# B&R Automation Studio project AS_Project (part 2)

#### Convert.c - dbGetData data conversion
```c
/********************************************************************
 * Library: AltDB
 * File: Convert.c
 ********************************************************************
 * dbGetData data conversion (Section 11). Converts the raw column
 * value bytes stored by Token.c (gConn[slot].ColValue[columnIdx])
 * into one of the DB_SQL_* target layouts of Table 22.
 *
 * Scope: the full conversion matrix (Table 23) is implemented for
 * the practically important source/target combinations. Combinations
 * marked '-' in Table 23, and sources this library cannot decode at
 * all (SQL_VARIANT, XML, UDT), are rejected with dbERR_DATABASE /
 * SQLSTATE 07006, matching the "not allowed" semantics of the
 * specification. DATETIMEOFFSET is read as if it were DATETIME2 (the
 * trailing minute-offset field is ignored, i.e. treated as UTC/local
 * time) - a documented simplification, see Common.h.
 ********************************************************************/
#include <bur/plctypes.h>
#include <runtime.h>
#include <AsTCP.h>
#include <AltDB.h>
#include "Common.h"
#include <string.h>

enum {
	FAM_INT, FAM_FLOAT, FAM_DECIMAL, FAM_MONEY, FAM_CHAR, FAM_BINARY,
	FAM_DATE, FAM_TIME, FAM_DATETIME, FAM_DATETIME2, FAM_GUID, FAM_UNSUPPORTED
};

static int Family(unsigned char t)
{
	switch (t) {
	case 0x30: case 0x32: case 0x34: case 0x38: case 0x7F:
	case 0x26: case 0x68:
		return FAM_INT;
	case 0x3B: case 0x3E: case 0x6D:
		return FAM_FLOAT;
	case 0x6A: case 0x6C:
		return FAM_DECIMAL;
	case 0x3C: case 0x7A: case 0x6E:
		return FAM_MONEY;
	case 0xA7: case 0xAF: case 0xE7: case 0xEF:
	case 0x2F: case 0x27:
	case 0x23: case 0x63:
		return FAM_CHAR;
	case 0xA5: case 0xAD: case 0x2D: case 0x25: case 0x22:
		return FAM_BINARY;
	case 0x28:
		return FAM_DATE;
	case 0x29:
		return FAM_TIME;
	case 0x3A: case 0x3D: case 0x6F:
		return FAM_DATETIME;
	case 0x2A: case 0x2B:
		return FAM_DATETIME2;
	case 0x24:
		return FAM_GUID;
	default:
		return FAM_UNSUPPORTED;
	}
}

static long long ReadIntValue(const unsigned char *p, UDINT len)
{
	unsigned long long u = 0;
	UDINT i;
	for (i = 0; i < len && i < 8; i++) u |= ((unsigned long long)p[i]) << (8 * i);
	if (len == 1) return (long long)u;        /* tinyint/bit: unsigned */
	if (len == 2) return (long long)(short)(unsigned short)u;
	if (len == 4) return (long long)(DINT)(UDINT)u;
	return (long long)u;
}

static long long ReadMoneyValue(const unsigned char *p, UDINT len)
{
	if (len == 4) return (long long)(DINT)AltDB_ReadLE32(p);
	{
		DINT hi = (DINT)AltDB_ReadLE32(p);
		UDINT lo = AltDB_ReadLE32(p + 4);
		return ((long long)hi << 32) | (long long)lo;
	}
}

static double ReadFloatValue(const unsigned char *p, UDINT len)
{
	if (len == 4) {
		union { UDINT u; float f; } v;
		v.u = AltDB_ReadLE32(p);
		return (double)v.f;
	} else {
		union { unsigned long long u; double d; } v;
		v.u = AltDB_ReadLE64(p);
		return v.d;
	}
}

/* value = integer / 10^scale, formatted as a decimal string */
static UDINT FormatScaledI64(long long v, USINT scale, char *dst, UDINT dstCap)
{
	unsigned char mag[8];
	BOOL positive = (v >= 0);
	unsigned long long u = positive ? (unsigned long long)v : (unsigned long long)(-(v + 1)) + 1ULL;
	UDINT i;
	for (i = 0; i < 8; i++) { mag[i] = (unsigned char)(u & 0xFF); u >>= 8; }
	return AltDB_FormatDecimal(mag, 8, positive, scale, dst, dstCap);
}

/* Decodes a DECIMALN/NUMERICN value (1 sign byte + little-endian
 * magnitude) into a plain double; sufficient precision for REAL /
 * DOUBLE targets (exact string output uses AltDB_FormatDecimal
 * directly for the CHAR target). */
static double DecimalToDouble(const unsigned char *raw, UDINT len, USINT scale)
{
	double v = 0.0;
	UDINT magLen = (len > 0) ? len - 1 : 0;
	BOOL positive = (len > 0) ? (raw[0] != 0) : TRUE;
	double divisor = 1.0;
	UDINT i;

	for (i = magLen; i > 0; i--) {
		v = v * 256.0 + (double)raw[i];
	}
	if (!positive) v = -v;
	for (i = 0; i < scale; i++) divisor *= 10.0;
	return v / divisor;
}

static void WriteGuidString(const unsigned char *g, char *dst)
{
	static const char *hex = "0123456789ABCDEF";
	static const int order[16] = {3,2,1,0, 5,4, 7,6, 8,9, 10,11,12,13,14,15};
	int i, p = 0;
	for (i = 0; i < 16; i++) {
		unsigned char b = g[order[i]];
		dst[p++] = hex[(b >> 4) & 0xF];
		dst[p++] = hex[b & 0xF];
		if (i == 3 || i == 5 || i == 7 || i == 9) dst[p++] = '-';
	}
	dst[p] = 0;
}

/* ---------------- date / time decoding (Section 10.9) ---------------- */

/* Howard Hinnant's civil_from_days algorithm (public domain formula),
 * valid over the whole proleptic Gregorian calendar. z = days since
 * 1970-01-01. */
static void CivilFromDays(long long z, INT *y, UINT *m, UINT *d)
{
	long long era;
	unsigned doe, yoe, doy, mp;

	z += 719468;
	era = (z >= 0 ? z : z - 146096) / 146097;
	doe = (unsigned)(z - era * 146097);
	yoe = (doe - doe / 1460 + doe / 36524 - doe / 146096) / 365;
	doy = doe - (365 * yoe + yoe / 4 - yoe / 100);
	mp = (5 * doy + 2) / 153;
	*d = (UINT)(doy - (153 * mp + 2) / 5 + 1);
	*m = (UINT)(mp + (mp < 10 ? 3 : -9));
	*y = (INT)((long long)yoe + era * 400 + (*m <= 2 ? 1 : 0));
}

typedef struct { INT y; UINT mo; UINT d; UINT h; UINT mi; UINT s; UDINT frac; USINT fracDigits; } DecodedDT;

/* days-since-0001-01-01 -> civil date */
static void DateFromDbDays(UDINT dbDays, INT *y, UINT *m, UINT *d)
{
	/* days_from_civil(1,1,1) = -719162 (date 0001-01-01 relative to 1970-01-01) */
	CivilFromDays((long long)dbDays - 719162LL, y, m, d);
}

static BOOL DecodeDateTime(int fam, unsigned char dataType, const unsigned char *raw, UDINT rawLen, USINT scale, DecodedDT *out)
{
	memset(out, 0, sizeof(*out));

	if (fam == FAM_DATE) {
		UDINT days = raw[0] | ((UDINT)raw[1] << 8) | ((UDINT)raw[2] << 16);
		DateFromDbDays(days, &out->y, &out->mo, &out->d);
		return TRUE;
	}
	if (fam == FAM_TIME || fam == FAM_DATETIME2) {
		UDINT dateBytes = (fam == FAM_DATETIME2) ? 3 : 0;
		UDINT offsetBytes = (dataType == 0x2B) ? 2 : 0;
		UDINT timeLen = (rawLen > dateBytes + offsetBytes) ? rawLen - dateBytes - offsetBytes : rawLen;
		UDINT i;
		unsigned long long ticks = 0;
		unsigned long long divisor = 1;
		UDINT secTotal;

		for (i = 0; i < timeLen && i < 8; i++) ticks |= ((unsigned long long)raw[i]) << (8 * i);
		for (i = 0; i < scale; i++) divisor *= 10ULL;
		secTotal = (UDINT)(ticks / divisor);
		out->frac = (UDINT)(ticks % divisor);
		out->fracDigits = scale;
		out->h = secTotal / 3600; out->mi = (secTotal / 60) % 60; out->s = secTotal % 60;

		if (fam == FAM_DATETIME2) {
			UDINT days = raw[timeLen] | ((UDINT)raw[timeLen + 1] << 8) | ((UDINT)raw[timeLen + 2] << 16);
			DateFromDbDays(days, &out->y, &out->mo, &out->d);
		}
		return TRUE;
	}
	if (fam == FAM_DATETIME) {
		if (rawLen == 4) { /* SMALLDATETIME: days(2,u16) + minutes(2,u16) since 1900-01-01 */
			UINT days = (UINT)AltDB_ReadLE16(raw);
			UINT minutes = (UINT)AltDB_ReadLE16(&raw[2]);
			CivilFromDays((long long)days - 25567LL, &out->y, &out->mo, &out->d); /* 1900-01-01 vs 1970-01-01 */
			out->h = minutes / 60; out->mi = minutes % 60; out->s = 0;
		} else { /* DATETIME: days(4,signed) + ticks(4,u32) of 1/300s since midnight */
			DINT days = (DINT)AltDB_ReadLE32(raw);
			UDINT ticks = AltDB_ReadLE32(&raw[4]);
			UDINT secTotal = ticks / 300;
			CivilFromDays((long long)days - 25567LL, &out->y, &out->mo, &out->d);
			out->h = secTotal / 3600; out->mi = (secTotal / 60) % 60; out->s = secTotal % 60;
		}
		return TRUE;
	}
	return FALSE;
}

static UDINT FormatDateTimeChar(int fam, const DecodedDT *dt, char *dst, UDINT cap)
{
	UDINT n = 0;
	char tmp[16];
	UDINT tn;

#define APPEND_NUM(v, width) do { \
		UDINT k; tn = (UDINT)AltDB_FormatI64((v), tmp, sizeof(tmp)); \
		for (k = tn; k < (UDINT)(width); k++) { if (n < cap) dst[n++] = '0'; } \
		for (k = 0; k < tn; k++) { if (n < cap) dst[n++] = tmp[k]; } \
	} while (0)

	if (fam == FAM_DATE || fam == FAM_DATETIME || fam == FAM_DATETIME2) {
		APPEND_NUM(dt->y, 4);
		if (n < cap) dst[n++] = '-';
		APPEND_NUM((long long)dt->mo, 2);
		if (n < cap) dst[n++] = '-';
		APPEND_NUM((long long)dt->d, 2);
		if (fam == FAM_DATE) { if (n < cap) dst[n] = 0; return n; }
		if (n < cap) dst[n++] = ' ';
	}

	APPEND_NUM((long long)dt->h, 2);
	if (n < cap) dst[n++] = ':';
	APPEND_NUM((long long)dt->mi, 2);
	if (n < cap) dst[n++] = ':';
	APPEND_NUM((long long)dt->s, 2);
	if (dt->fracDigits > 0) {
		if (n < cap) dst[n++] = '.';
		APPEND_NUM((long long)dt->frac, dt->fracDigits);
	}
	if (n < cap) dst[n] = 0;
	return n;
#undef APPEND_NUM
}

static void PutCharResult(const char *text, UDINT textLen, UDINT pData, UDINT dataSize,
                           UINT *status, INT *dbError, UDINT *actDataSize)
{
	UDINT required = textLen + 1;
	if (dataSize < required) {
		*status = dbERR_BUFFER_SIZE; *dbError = DB_SQL_ERROR; *actDataSize = required;
		return;
	}
	memcpy((void *)pData, text, textLen);
	((char *)pData)[textLen] = 0;
	*status = ERR_OK; *dbError = 0; *actDataSize = required;
}

void AltDB_GetData(UDINT slot, UDINT columnIdx, INT dataType, UDINT pData, UDINT dataSize,
                      UINT *status, INT *dbError, UDINT *actDataSize)
{
	ConnSlot *c = &gConn[slot];
	UDINT idx;
	ColumnInfo *col;
	int fam;
	const unsigned char *raw;
	UDINT rawLen;

	*actDataSize = 0;

	if (!c->RowReady) { *status = dbERR_SQL_EXECUTE_REQUIRED; *dbError = DB_SQL_ERROR; return; }
	if (columnIdx == 0 || columnIdx > (UDINT)c->ColumnCount || columnIdx > ND_MAX_COLUMNS) {
		*status = dbERR_INVALID_COLUMN; *dbError = DB_SQL_ERROR; return;
	}
	if (pData == 0) { *status = dbERR_NULLPOINTER; *dbError = DB_SQL_ERROR; return; }

	idx = columnIdx - 1;
	if (c->ColAlreadyRead[idx]) { *status = dbERR_DATABASE; *dbError = DB_SQL_NO_DATA; return; }

	if (c->ColIsNull[idx]) {
		*status = ERR_OK; *dbError = 0; *actDataSize = 0xFFFFFFFFUL;
		c->ColAlreadyRead[idx] = TRUE;
		return;
	}

	col = &c->Columns[idx];
	raw = c->ColValue[idx];
	rawLen = c->ColValueLen[idx];
	if (rawLen > ND_MAX_COL_VALUE_LEN) rawLen = ND_MAX_COL_VALUE_LEN;

	if (!col->Supported) {
		AltDB_DiagPushClient(slot, "07006", "source column type is not convertible by this library");
		*status = dbERR_DATABASE; *dbError = DB_SQL_ERROR; return;
	}

	fam = Family(col->DataType);

	switch (dataType) {

	case 1: { /* DB_SQL_CHAR */
		char text[600];
		UDINT n = 0;

		switch (fam) {
		case FAM_CHAR:
			if (col->IsUnicode) n = AltDB_WireToConn(c->Encoding, raw, rawLen, (unsigned char *)text, sizeof(text) - 1);
			else { n = (rawLen < sizeof(text) - 1) ? rawLen : sizeof(text) - 1; memcpy(text, raw, n); }
			break;
		case FAM_BINARY: {
			static const char *hex = "0123456789ABCDEF";
			UDINT i;
			for (i = 0; i < rawLen && n + 2 < sizeof(text); i++) {
				text[n++] = hex[(raw[i] >> 4) & 0xF];
				text[n++] = hex[raw[i] & 0xF];
			}
			break;
		}
		case FAM_INT:
			n = (UDINT)AltDB_FormatI64(ReadIntValue(raw, rawLen), text, sizeof(text));
			break;
		case FAM_MONEY:
			n = FormatScaledI64(ReadMoneyValue(raw, rawLen), 4, text, sizeof(text));
			break;
		case FAM_DECIMAL:
			n = AltDB_FormatDecimal(&raw[1], (rawLen > 0) ? rawLen - 1 : 0, raw[0] != 0, col->Scale, text, sizeof(text));
			break;
		case FAM_FLOAT:
			n = AltDB_FormatDouble(ReadFloatValue(raw, rawLen), (rawLen == 4) ? 7 : 15, text, sizeof(text));
			break;
		case FAM_GUID:
			if (rawLen >= 16) { WriteGuidString(raw, text); n = (UDINT)strlen(text); }
			break;
		case FAM_DATE: case FAM_TIME: case FAM_DATETIME: case FAM_DATETIME2: {
			DecodedDT dt;
			if (DecodeDateTime(fam, col->DataType, raw, rawLen, col->Scale, &dt)) {
				n = FormatDateTimeChar(fam, &dt, text, sizeof(text));
			}
			break;
		}
		default:
			AltDB_DiagPushClient(slot, "07006", "source column type is not convertible to DB_SQL_CHAR");
			*status = dbERR_DATABASE; *dbError = DB_SQL_ERROR; return;
		}
		PutCharResult(text, n, pData, dataSize, status, dbError, actDataSize);
		if (*status == ERR_OK) c->ColAlreadyRead[idx] = TRUE;
		return;
	}

	case -6: case 5: case 4: case -25: { /* TINYINT / SMALLINT / INTEGER / BIGINT */
		long long v;
		UDINT needed = (dataType == -6) ? 1 : (dataType == 5) ? 2 : (dataType == 4) ? 4 : 8;

		if (fam == FAM_INT) v = ReadIntValue(raw, rawLen);
		else if (fam == FAM_MONEY) v = ReadMoneyValue(raw, rawLen) / 10000;
		else if (fam == FAM_DECIMAL) v = (long long)DecimalToDouble(raw, rawLen, col->Scale);
		else if (fam == FAM_FLOAT) v = (long long)ReadFloatValue(raw, rawLen);
		else {
			AltDB_DiagPushClient(slot, "07006", "source column type is not convertible to an integer type");
			*status = dbERR_DATABASE; *dbError = DB_SQL_ERROR; return;
		}
				/* AsDB compatibility: allow BIGINT -> UDINT */

		if (dataType == -25 && dataSize == 4)
		{
			UDINT tmp = (UDINT)v;
			memcpy((void *)pData, &tmp, 4);
			*status = ERR_OK;
			*dbError = 0;
			*actDataSize = 4;
			c->ColAlreadyRead[idx] = TRUE;
			return;
		}
		if (dataSize < needed) { *status = dbERR_BUFFER_SIZE; *dbError = DB_SQL_ERROR; *actDataSize = needed; return; }
		{
			unsigned char tmp[8];
			UDINT i;
			for (i = 0; i < needed; i++) tmp[i] = (unsigned char)((unsigned long long)v >> (8 * i));
			memcpy((void *)pData, tmp, needed);
		}
		*status = ERR_OK; *dbError = 0; *actDataSize = needed;
		c->ColAlreadyRead[idx] = TRUE;
		return;
	}

	case 7: case 8: { /* DB_SQL_REAL / DB_SQL_DOUBLE */
		double v;
		UDINT needed = (dataType == 7) ? 4 : 8;

		if (fam == FAM_INT) v = (double)ReadIntValue(raw, rawLen);
		else if (fam == FAM_MONEY) v = (double)ReadMoneyValue(raw, rawLen) / 10000.0;
		else if (fam == FAM_DECIMAL) v = DecimalToDouble(raw, rawLen, col->Scale);
		else if (fam == FAM_FLOAT) v = ReadFloatValue(raw, rawLen);
		else {
			AltDB_DiagPushClient(slot, "07006", "source column type is not convertible to a floating point type");
			*status = dbERR_DATABASE; *dbError = DB_SQL_ERROR; return;
		}
		if (dataSize < needed) { *status = dbERR_BUFFER_SIZE; *dbError = DB_SQL_ERROR; *actDataSize = needed; return; }
		if (needed == 4) {
			union { UDINT u; float f; } u; u.f = (float)v;
			memcpy((void *)pData, &u.u, 4);
		} else {
			union { unsigned long long u; double d; } u; u.d = v;
			memcpy((void *)pData, &u.u, 8);
		}
		*status = ERR_OK; *dbError = 0; *actDataSize = needed;
		c->ColAlreadyRead[idx] = TRUE;
		return;
	}

	case 9: case 10: case 11: { /* DB_SQL_DATE / DB_SQL_TIME / DB_SQL_TIMESTAMP */
		DecodedDT dt;
		UDINT needed = (dataType == 9 || dataType == 10) ? 6 : 12;
		UINT vals[6];

		if (fam != FAM_DATE && fam != FAM_TIME && fam != FAM_DATETIME && fam != FAM_DATETIME2) {
			AltDB_DiagPushClient(slot, "07006", "source column type is not convertible to a date/time type");
			*status = dbERR_DATABASE; *dbError = DB_SQL_ERROR; return;
		}
		if (dataType == 9 && fam == FAM_TIME) {
			AltDB_DiagPushClient(slot, "07006", "TIME source cannot convert to DB_SQL_DATE");
			*status = dbERR_DATABASE; *dbError = DB_SQL_ERROR; return;
		}
		if (!DecodeDateTime(fam, col->DataType, raw, rawLen, col->Scale, &dt)) {
			*status = dbERR_DATABASE; *dbError = DB_SQL_ERROR; return;
		}
		if (dataSize < needed) { *status = dbERR_BUFFER_SIZE; *dbError = DB_SQL_ERROR; *actDataSize = needed; return; }

		if (dataType == 9) { vals[0] = (UINT)dt.y; vals[1] = dt.mo; vals[2] = dt.d; }
		else if (dataType == 10) { vals[0] = dt.h; vals[1] = dt.mi; vals[2] = dt.s; }
		else { vals[0] = (UINT)dt.y; vals[1] = dt.mo; vals[2] = dt.d; vals[3] = dt.h; vals[4] = dt.mi; vals[5] = dt.s; }
		{
			UDINT n = (dataType == 11) ? 6 : 3;
			UDINT i;
			for (i = 0; i < n; i++) AltDB_WriteLE16((unsigned char *)pData + i * 2, vals[i]);
		}
		*status = ERR_OK; *dbError = 0; *actDataSize = needed;
		c->ColAlreadyRead[idx] = TRUE;
		return;
	}

	case -11: { /* DB_SQL_GUID */
		if (fam != FAM_GUID && !(fam == FAM_BINARY && rawLen == 16)) {
			AltDB_DiagPushClient(slot, "07006", "source column type is not convertible to DB_SQL_GUID");
			*status = dbERR_DATABASE; *dbError = DB_SQL_ERROR; return;
		}
		if (dataSize < 16) { *status = dbERR_BUFFER_SIZE; *dbError = DB_SQL_ERROR; *actDataSize = 16; return; }
		memcpy((void *)pData, raw, 16);
		*status = ERR_OK; *dbError = 0; *actDataSize = 16;
		c->ColAlreadyRead[idx] = TRUE;
		return;
	}

	case 2: case 3: { /* DB_SQL_NUMERIC / DB_SQL_DECIMAL: ODBC SQL_NUMERIC_STRUCT (19 bytes) */
		unsigned char prec, scale, sign;
		unsigned char val[16];

		memset(val, 0, sizeof(val));
		if (fam == FAM_DECIMAL) {
			UDINT magLen = (rawLen > 0) ? rawLen - 1 : 0;
			if (magLen > 16) magLen = 16;
			memcpy(val, &raw[1], magLen);
			sign = (raw[0] != 0) ? 1 : 0;
			prec = col->Precision; scale = col->Scale;
		} else if (fam == FAM_INT || fam == FAM_MONEY) {
			long long v = (fam == FAM_INT) ? ReadIntValue(raw, rawLen) : ReadMoneyValue(raw, rawLen);
			unsigned long long u = (v >= 0) ? (unsigned long long)v : (unsigned long long)(-(v + 1)) + 1ULL;
			UDINT i;
			for (i = 0; i < 8; i++) { val[i] = (unsigned char)(u & 0xFF); u >>= 8; }
			sign = (v >= 0) ? 1 : 0;
			scale = (fam == FAM_MONEY) ? 4 : 0;
			prec = 19;
		} else {
			AltDB_DiagPushClient(slot, "07006", "source column type is not convertible to DB_SQL_NUMERIC/DECIMAL");
			*status = dbERR_DATABASE; *dbError = DB_SQL_ERROR; return;
		}
		if (dataSize < 19) { *status = dbERR_BUFFER_SIZE; *dbError = DB_SQL_ERROR; *actDataSize = 19; return; }
		{
			unsigned char *out = (unsigned char *)pData;
			out[0] = prec; out[1] = (unsigned char)scale; out[2] = sign;
			memcpy(&out[3], val, 16);
		}
		*status = ERR_OK; *dbError = 0; *actDataSize = 19;
		c->ColAlreadyRead[idx] = TRUE;
		return;
	}

	default:
		AltDB_DiagPushClient(slot, "HY004", "unsupported dataType requested");
		*status = dbERR_INVALID_DATATYPE; *dbError = DB_SQL_ERROR;
		return;
	}
}
```

#### Connect.c - dbConnect, dbConnectEnc
```c
/********************************************************************
 * Library: AltDB
 * File: Connect.c
 ********************************************************************
 * dbConnect / dbConnectEnc (Section 7.2-7.4).
 ********************************************************************/
#include <bur/plctypes.h>
#include <runtime.h>
#include <AsTCP.h>
#include <AltDB.h>
#include "Common.h"
#include <string.h>

static BOOL EqualsIgnoreCase(const char *a, const char *b)
{
	while (*a && *b) {
		char ca = *a, cb = *b;
		if (ca >= 'a' && ca <= 'z') ca = (char)(ca - 'a' + 'A');
		if (cb >= 'a' && cb <= 'z') cb = (char)(cb - 'a' + 'A');
		if (ca != cb) return FALSE;
		a++; b++;
	}
	return (*a == 0 && *b == 0);
}

/* Parsed/validated dbConnect/dbConnectEnc inputs, independent of any
 * connection slot (no slot is needed just to validate). */
typedef struct ParsedConnectInputs
{
	char   hostBuf[128];	/* NUL-terminated, port and named-instance suffix stripped */
	UDINT  hostLen;
	UINT   port;
	UINT   encoding;		/* DBENC_ISO_8859_1 / DBENC_UTF_8 */
	const char *user;
	UDINT  userLen;
	const char *pass;
	UDINT  passLen;
	const char *db;
	UDINT  dbLen;
} ParsedConnectInputs;

/* Validates dbConnect/dbConnectEnc inputs and fills *out. Performs no
 * slot allocation or lookup, so the caller can validate (cheap) before
 * committing to a slot allocation or lock (preserves AsDb's original
 * error precedence, e.g. an unsupported databaseSystem is reported
 * even when the connection pool happens to be full). On failure,
 * status and dbError are set and *out is left in an undefined state. */
static BOOL ValidateAndParseConnectInputs(UDINT pServerName, UDINT pUserName, UDINT pPassword,
	UDINT pDatabaseName, UDINT databaseSystem, UDINT pEncoding,
	ParsedConnectInputs *out, UINT *status, INT *dbError)
{
	const char *server = (const char *)pServerName;
	const char *colon;
	const char *backslash;
	char hostPortBuf[128];
	UDINT hostPortLen;

	if (databaseSystem != DB_SYSTEM_MS_SQL) {
		*status = dbERR_UNSUPPORTED_DATABASE; *dbError = DB_SQL_ERROR; return FALSE;
	}
	if (pServerName == 0 || pUserName == 0 || pPassword == 0 || pDatabaseName == 0) {
		*status = dbERR_NULLPOINTER; *dbError = DB_SQL_ERROR; return FALSE;
	}
	out->user = (const char *)pUserName;
	out->pass = (const char *)pPassword;
	out->db = (const char *)pDatabaseName;
	out->userLen = (UDINT)strlen(out->user);
	out->passLen = (UDINT)strlen(out->pass);
	out->dbLen = (UDINT)strlen(out->db);

	if (out->userLen > 128) { *status = dbERR_INVALID_USERNAME; *dbError = DB_SQL_ERROR; return FALSE; }
	if (out->passLen > 128) { *status = dbERR_INVALID_PASSWORD; *dbError = DB_SQL_ERROR; return FALSE; }
	if (out->dbLen < 1 || out->dbLen > 128) {
		*status = dbERR_INVALID_DATABASE_NAME; *dbError = DB_SQL_ERROR; return FALSE;
	}

	/* Strip an optional backslash-prefixed instance-name suffix (SQL
	 * Server named-instance syntax, e.g. "192.168.66.99:1433" followed
	 * by "SQLEXPRESS"). Named-instance resolution via the SQL Server
	 * Browser service (UDP 1434) is out of scope for this library,
	 * exactly as for the original AsDb (a fixed TCP port is required
	 * either way), so the instance name is accepted for drop-in
	 * compatibility but otherwise ignored; only the host[:port] part
	 * before the backslash is parsed and used to connect. */
	backslash = strchr(server, '\\');
	hostPortLen = backslash ? (UDINT)(backslash - server) : (UDINT)strlen(server);
	if (hostPortLen == 0 || hostPortLen > sizeof(hostPortBuf) - 1) {
		*status = dbERR_INVALID_SERVERNAME; *dbError = DB_SQL_ERROR; return FALSE;
	}
	memcpy(hostPortBuf, server, hostPortLen); hostPortBuf[hostPortLen] = 0;

	colon = strrchr(hostPortBuf, ':');
	if (colon != NULL) {
		long p = 0;
		UDINT i;
		BOOL okDigits = (colon[1] != 0);
		for (i = 0; colon[1 + i] != 0; i++) {
			char ch = colon[1 + i];
			if (ch < '0' || ch > '9') { okDigits = FALSE; break; }
			p = p * 10 + (ch - '0');
		}
		out->hostLen = (UDINT)(colon - hostPortBuf);
		if (!okDigits || p < 1 || p > 65535 || out->hostLen == 0) {
			*status = dbERR_INVALID_SERVERNAME; *dbError = DB_SQL_ERROR; return FALSE;
		}
		out->port = (UINT)p;
	} else {
		out->hostLen = (UDINT)strlen(hostPortBuf);
		if (out->hostLen == 0) {
			*status = dbERR_INVALID_SERVERNAME; *dbError = DB_SQL_ERROR; return FALSE;
		}
		out->port = 1433; /* default MS SQL port, [V-03] */
	}
	memcpy(out->hostBuf, hostPortBuf, out->hostLen); out->hostBuf[out->hostLen] = 0;

	out->encoding = DBENC_ISO_8859_1;
	if (pEncoding != 0) {
		const char *enc = (const char *)pEncoding;
		if (EqualsIgnoreCase(enc, "UTF-8")) out->encoding = DBENC_UTF_8;
		else if (EqualsIgnoreCase(enc, "ISO-8859-1")) out->encoding = DBENC_ISO_8859_1;
		else {
			*status = dbERR_UNSUPPORTED_ENCODING; *dbError = DB_SQL_ERROR; return FALSE;
		}
	}

	return TRUE;
}

/* Copies already-validated inputs into the slot's login parameters.
 * Shared by (a) the first allocation of a new connection and (b)
 * re-capturing possibly-corrected inputs after a connect job was
 * abandoned via enable := FALSE while still in progress (Section 9.3
 * job cancellation; see CustomerChangeAnalysis.md item 1). */
static void CommitConnectInputsToSlot(UDINT slot, const ParsedConnectInputs *in)
{
	gConn[slot].Encoding = in->encoding;
	memcpy(gConn[slot].HostBuf, in->hostBuf, in->hostLen + 1);
	gConn[slot].Port = in->port;
	gConn[slot].LoginUserLen = in->userLen;
	memcpy(gConn[slot].LoginUser, in->user, in->userLen + 1);
	gConn[slot].LoginPassLen = in->passLen;
	memcpy(gConn[slot].LoginPass, in->pass, in->passLen + 1);
	gConn[slot].LoginDbLen = in->dbLen;
	memcpy(gConn[slot].LoginDb, in->db, in->dbLen + 1);
}

static void ConnectCommon(UDINT instAddr, BOOL enable, UDINT pServerName, UDINT pUserName, UDINT pPassword,
	UDINT pDatabaseName, UDINT databaseSystem, UDINT pEncoding,
	UINT *status, INT *dbError, UDINT *connectionIdent)
{
	UDINT slot;
	UINT generation;
	INT r;

	if (!enable) {
		if (*connectionIdent != 0 && AltDB_SlotFromHandle(*connectionIdent, &slot, &generation) &&
		AltDB_IsOwner(slot, instAddr)) {
			/* Tear down the in-flight connection instead of leaving a
			 * half-finished handshake (and a leaked TCP socket) behind.
			 * Best-effort and non-blocking: if the close needs more
			 * cycles than this single call, it is completed either by
			 * a later enable := FALSE call on this same instance or by
			 * the Abandoned-recapture path below on the next
			 * dbConnect/dbConnectEnc call for this handle. */
			AltDB_NetDisconnectStep(slot);
			gConn[slot].Abandoned = TRUE;
			AltDB_Unlock(slot);
		}
		*status = ERR_FUB_ENABLE_FALSE; *dbError = 0;
		return;
	}

	if (*connectionIdent == 0) {
		ParsedConnectInputs parsed;

		if (!ValidateAndParseConnectInputs(pServerName, pUserName, pPassword, pDatabaseName,
		databaseSystem, pEncoding, &parsed, status, dbError)) {
			return; /* no slot allocated yet, nothing to release */
		}
		if (!AltDB_SlotAlloc(&slot)) { *status = dbERR_MEMORY; *dbError = DB_SQL_ERROR; return; }
		generation = gConn[slot].Generation;

		CommitConnectInputsToSlot(slot, &parsed);
		gConn[slot].JobKind = JOB_CONNECT;
		gConn[slot].State = CONNSTATE_OPENING;
		AltDB_DiagClear(slot);

		*connectionIdent = AltDB_MakeHandle(slot, generation);
	} else {
		if (!AltDB_SlotFromHandle(*connectionIdent, &slot, &generation)) {
			*status = dbERR_DATABASE; *dbError = DB_SQL_ERROR; return;
		}

		if (gConn[slot].Abandoned) {
			/* Previous connect job on this handle was cancelled
			 * mid-flight (enable := FALSE while BUSY). Re-validate and
			 * re-capture the current inputs (the application may have
			 * corrected them, e.g. the password) before touching the
			 * lock, then finish closing any socket left over from the
			 * abandoned attempt and restart the handshake from
			 * CONNSTATE_OPENING rather than blindly resuming stale
			 * state. */
			ParsedConnectInputs parsed;

			if (!ValidateAndParseConnectInputs(pServerName, pUserName, pPassword, pDatabaseName,
			databaseSystem, pEncoding, &parsed, status, dbError)) {
				return; /* still Abandoned, lock untouched; caller may retry */
			}
			if (!AltDB_TryLock(slot, instAddr)) { *status = ERR_FUB_BUSY; return; }
			if (AltDB_NetDisconnectStep(slot) == NET_IN_PROGRESS) {
				*status = ERR_FUB_BUSY; return; /* lock held; finish closing on the next call */
			}
			CommitConnectInputsToSlot(slot, &parsed);
			gConn[slot].Abandoned = FALSE;
			gConn[slot].JobKind = JOB_CONNECT;
			gConn[slot].State = CONNSTATE_OPENING;
			AltDB_DiagClear(slot);
		} else if (gConn[slot].JobKind != JOB_CONNECT) {
			*status = dbERR_DATABASE; *dbError = DB_SQL_ERROR; return;
		}
	}

	if (!AltDB_TryLock(slot, instAddr)) { *status = ERR_FUB_BUSY; return; }

	r = AltDB_NetConnectStep(slot);
	if (r == NET_IN_PROGRESS) { *status = ERR_FUB_BUSY; return; }

	AltDB_Unlock(slot);
	if (r == NET_DONE) {
		*status = ERR_OK;
		*dbError = 0;
	} else {
		*status = dbERR_DATABASE;
		*dbError = DB_SQL_ERROR;
	}
}

void dbConnect(struct dbConnect *inst)
{
	ConnectCommon((UDINT)inst, inst->enable, inst->pServerName, inst->pUserName, inst->pPassword,
		inst->pDatabaseName, inst->databaseSystem, 0,
		&inst->status, &inst->dbError, &inst->connectionIdent);
}

void dbConnectEnc(struct dbConnectEnc *inst)
{
	ConnectCommon((UDINT)inst, inst->enable, inst->pServerName, inst->pUserName, inst->pPassword,
		inst->pDatabaseName, inst->databaseSystem, inst->pEncoding,
		&inst->status, &inst->dbError, &inst->connectionIdent);
}
```

#### Execute.c - dbExecuteSql, dbGetAffectedRows, dbGetColumnCount
```c
/********************************************************************
 * Library: AltDB
 * File: Execute.c
 ********************************************************************
 * dbExecuteSql (Section 7.5), dbGetAffectedRows (7.6),
 * dbGetColumnCount (7.7).
 ********************************************************************/
#include <bur/plctypes.h>
#include <runtime.h>
#include <AsTCP.h>
#include <AltDB.h>
#include "Common.h"
#include <string.h>

#define EXECSTEP_DRAIN 0
#define EXECSTEP_SEND  1
#define EXECSTEP_RECV  2

static BOOL IsBrokenState(UINT state)
{
	return (state == CONNSTATE_BROKEN || state == CONNSTATE_FAILED);
}

void dbExecuteSql(struct dbExecuteSql *inst)
{
	UDINT instAddr = (UDINT)inst;
	UDINT slot;
	UINT generation;
	BOOL fresh;

	if (!inst->enable) {
		if (AltDB_SlotFromHandle(inst->connectionIdent, &slot, &generation) && AltDB_IsOwner(slot, instAddr)) {
			AltDB_Unlock(slot);
		}
		inst->status = ERR_FUB_ENABLE_FALSE; inst->dbError = 0;
		return;
	}

	if (!AltDB_SlotFromHandle(inst->connectionIdent, &slot, &generation)) {
		inst->status = dbERR_INVALID_HANDLE; inst->dbError = DB_SQL_INVALID_HANDLE; return;
	}
	if (IsBrokenState(gConn[slot].State)) {
		AltDB_DiagPushClient(slot, "08S01", "connection is broken, call dbDisconnect");
		inst->status = dbERR_DATABASE; inst->dbError = DB_SQL_ERROR; return;
	}

	fresh = !gConn[slot].Locked;
	if (!fresh) {
		if (gConn[slot].JobOwner != instAddr) { inst->status = ERR_FUB_BUSY; return; }
		if (gConn[slot].JobKind != JOB_EXECUTE) {
			AltDB_DiagPushClient(slot, "HY010", "function sequence error");
			inst->status = dbERR_DATABASE; inst->dbError = DB_SQL_ERROR; return;
		}
	}

	if (fresh) {
		const char *sql;
		UDINT sqlLen;

		if (!AltDB_TryLock(slot, instAddr)) { inst->status = ERR_FUB_BUSY; return; }
		gConn[slot].JobKind = JOB_EXECUTE;

		sql = (const char *)inst->pSqlStatement;
		if (inst->pSqlStatement == 0 || sql[0] == 0) {
			AltDB_Unlock(slot);
			inst->status = dbERR_INVALID_SQL_STATEMENT; inst->dbError = DB_SQL_ERROR; return;
		}
		sqlLen = (UDINT)strlen(sql);
		if (sqlLen > SQL_MAX_LEN) {
			AltDB_Unlock(slot);
			inst->status = dbERR_INVALID_SQL_STATEMENT; inst->dbError = DB_SQL_ERROR; return;
		}

		AltDB_BuildSqlBatch(slot, sql, sqlLen);
		gConn[slot].NetStep = gConn[slot].ResultSetOpen ? EXECSTEP_DRAIN : EXECSTEP_SEND;
	}

	if (gConn[slot].NetStep == EXECSTEP_DRAIN) {
		INT pumped = AltDB_NetRecvPump(slot);
		INT tok;

		if (pumped < 0) {
			AltDB_Unlock(slot); gConn[slot].State = CONNSTATE_BROKEN;
			inst->status = dbERR_DATABASE; inst->dbError = DB_SQL_ERROR; return;
		}
		tok = AltDB_TokenStep(slot, TOKMODE_DRAIN);
		if (tok == TOK_NEED_MORE) { inst->status = ERR_FUB_BUSY; return; }
		/* whether drain ended cleanly or hit an error, the stale result
		 * is considered discarded either way (best-effort, Common.h) */
		gConn[slot].ResultSetOpen = FALSE;
		gConn[slot].NetStep = EXECSTEP_SEND;
		inst->status = ERR_FUB_BUSY;
		return;
	}

	if (gConn[slot].NetStep == EXECSTEP_SEND) {
		INT r = AltDB_NetSendStep(slot);

		if (r == NET_ERROR) {
			AltDB_Unlock(slot); gConn[slot].State = CONNSTATE_BROKEN;
			inst->status = dbERR_DATABASE; inst->dbError = DB_SQL_ERROR; return;
		}
		if (r == NET_DONE) {
			AltDB_DiagClear(slot);
			gConn[slot].ColumnCount = 0;
			gConn[slot].HasResultSet = FALSE;
			gConn[slot].ResultSetOpen = FALSE;
			gConn[slot].AffectedRows = 0;
			gConn[slot].AffectedRowsKnown = FALSE;
			gConn[slot].RowReady = FALSE;
			gConn[slot].NoMoreRows = FALSE;
			gConn[slot].RowOverflow = FALSE;
			gConn[slot].NetStep = EXECSTEP_RECV;
		}
		inst->status = ERR_FUB_BUSY;
		return;
	}

	/* EXECSTEP_RECV */
	{
		INT pumped = AltDB_NetRecvPump(slot);
		INT tok;

		if (pumped < 0) {
			AltDB_Unlock(slot); gConn[slot].State = CONNSTATE_BROKEN;
			inst->status = dbERR_DATABASE; inst->dbError = DB_SQL_ERROR; return;
		}
		tok = AltDB_TokenStep(slot, TOKMODE_EXEC);
		switch (tok) {
		case TOK_NEED_MORE:
			inst->status = ERR_FUB_BUSY;
			return;
		case TOK_GOT_COLMETADATA:
		case TOK_GOT_DONE_FINAL:
			AltDB_Unlock(slot);
			gConn[slot].StatementActive = TRUE;
			inst->status = ERR_OK;
			inst->dbError = (gConn[slot].DiagCount > 0) ? 1 : 0;
			return;
		case TOK_ERROR_MEMORY:
			AltDB_Unlock(slot);
			inst->status = dbERR_MEMORY; inst->dbError = DB_SQL_ERROR;
			return;
		default: /* TOK_ERROR */
			AltDB_Unlock(slot);
			inst->status = dbERR_DATABASE; inst->dbError = DB_SQL_ERROR;
			return;
		}
	}
}

void dbGetAffectedRows(struct dbGetAffectedRows *inst)
{
	UDINT instAddr = (UDINT)inst;
	UDINT slot;
	UINT generation;

	if (!inst->enable) { inst->status = ERR_FUB_ENABLE_FALSE; inst->dbError = 0; return; }
	if (!AltDB_SlotFromHandle(inst->connectionIdent, &slot, &generation)) {
		inst->status = dbERR_INVALID_HANDLE; inst->dbError = DB_SQL_INVALID_HANDLE; return;
	}
	if (gConn[slot].Locked && gConn[slot].JobOwner != instAddr) { inst->status = ERR_FUB_BUSY; return; }
	if (!gConn[slot].StatementActive) {
		inst->status = dbERR_SQL_EXECUTE_REQUIRED; inst->dbError = DB_SQL_ERROR; return;
	}
	if (gConn[slot].HasResultSet) {
		 inst->status = ERR_OK; inst->dbError = 0; inst->affectedRows = 0xFFFFFFFF; return;
	}
	inst->status = ERR_OK; inst->dbError = 0;
	inst->affectedRows = gConn[slot].AffectedRowsKnown ? gConn[slot].AffectedRows : 0;
}

void dbGetColumnCount(struct dbGetColumnCount *inst)
{
	UDINT instAddr = (UDINT)inst;
	UDINT slot;
	UINT generation;

	if (!inst->enable) { inst->status = ERR_FUB_ENABLE_FALSE; inst->dbError = 0; return; }
	if (!AltDB_SlotFromHandle(inst->connectionIdent, &slot, &generation)) {
		inst->status = dbERR_INVALID_HANDLE; inst->dbError = DB_SQL_INVALID_HANDLE; return;
	}
	if (gConn[slot].Locked && gConn[slot].JobOwner != instAddr) { inst->status = ERR_FUB_BUSY; return; }
	if (!gConn[slot].StatementActive) {
		inst->status = dbERR_SQL_EXECUTE_REQUIRED; inst->dbError = DB_SQL_ERROR; return;
	}
	inst->status = ERR_OK; inst->dbError = 0;
	inst->columnCount = gConn[slot].HasResultSet ? (INT)gConn[slot].ColumnCount : 0;
}
```

#### Fetch.c - dbFetchNextRow, dbGetData
```c
/********************************************************************
 * Library: AltDB
 * File: Fetch.c
 ********************************************************************
 * dbFetchNextRow (Section 7.8), dbGetData (7.9).
 ********************************************************************/
#include <bur/plctypes.h>
#include <runtime.h>
#include <AsTCP.h>
#include <AltDB.h>
#include "Common.h"

static BOOL IsBrokenState(UINT state)
{
	return (state == CONNSTATE_BROKEN || state == CONNSTATE_FAILED);
}

void dbFetchNextRow(struct dbFetchNextRow *inst)
{
	UDINT instAddr = (UDINT)inst;
	UDINT slot;
	UINT generation;
	BOOL fresh;

	if (!inst->enable) {
		if (AltDB_SlotFromHandle(inst->connectionIdent, &slot, &generation) && AltDB_IsOwner(slot, instAddr)) {
			AltDB_Unlock(slot);
		}
		inst->status = ERR_FUB_ENABLE_FALSE; inst->dbError = 0;
		return;
	}

	if (!AltDB_SlotFromHandle(inst->connectionIdent, &slot, &generation)) {
		inst->status = dbERR_INVALID_HANDLE; inst->dbError = DB_SQL_INVALID_HANDLE; return;
	}
	if (IsBrokenState(gConn[slot].State)) {
		AltDB_DiagPushClient(slot, "08S01", "connection is broken, call dbDisconnect");
		inst->status = dbERR_DATABASE; inst->dbError = DB_SQL_ERROR; return;
	}

	fresh = !gConn[slot].Locked;
	if (!fresh) {
		if (gConn[slot].JobOwner != instAddr) { inst->status = ERR_FUB_BUSY; return; }
		if (gConn[slot].JobKind != JOB_FETCH) {
			AltDB_DiagPushClient(slot, "HY010", "function sequence error");
			inst->status = dbERR_DATABASE; inst->dbError = DB_SQL_ERROR; return;
		}
	}

	if (fresh) {
		if (!AltDB_TryLock(slot, instAddr)) { inst->status = ERR_FUB_BUSY; return; }
		gConn[slot].JobKind = JOB_FETCH;
	}

	if (!gConn[slot].ResultSetOpen) {
		/* end of result set, or no SELECT result ever opened - the
		 * default AsDb end-of-data signalling [V-04] */
		AltDB_Unlock(slot);
		inst->status = dbERR_DATABASE; inst->dbError = DB_SQL_NO_DATA;
		return;
	}

	{
		INT pumped = AltDB_NetRecvPump(slot);
		INT tok;

		if (pumped < 0) {
			AltDB_Unlock(slot); gConn[slot].State = CONNSTATE_BROKEN;
			inst->status = dbERR_DATABASE; inst->dbError = DB_SQL_ERROR; return;
		}
		tok = AltDB_TokenStep(slot, TOKMODE_FETCH);
		switch (tok) {
		case TOK_NEED_MORE:
			inst->status = ERR_FUB_BUSY;
			return;
		case TOK_GOT_ROW:
			AltDB_Unlock(slot);
			inst->status = ERR_OK; inst->dbError = 0;
			return;
		case TOK_GOT_EOF:
			AltDB_Unlock(slot);
			inst->status = dbERR_DATABASE; inst->dbError = DB_SQL_NO_DATA;
			return;
		case TOK_ERROR_MEMORY:
			gConn[slot].ResultSetOpen = FALSE;
			gConn[slot].NoMoreRows = TRUE;
			AltDB_Unlock(slot);
			inst->status = dbERR_MEMORY; inst->dbError = DB_SQL_ERROR;
			return;
		default: /* TOK_ERROR */
			AltDB_Unlock(slot);
			inst->status = dbERR_DATABASE; inst->dbError = DB_SQL_ERROR;
			return;
		}
	}
}

void dbGetData(struct dbGetData *inst)
{
	UDINT instAddr = (UDINT)inst;
	UDINT slot;
	UINT generation;

	if (!inst->enable) { inst->status = ERR_FUB_ENABLE_FALSE; inst->dbError = 0; return; }
	if (!AltDB_SlotFromHandle(inst->connectionIdent, &slot, &generation)) {
		inst->status = dbERR_INVALID_HANDLE; inst->dbError = DB_SQL_INVALID_HANDLE; return;
	}
	if (gConn[slot].Locked && gConn[slot].JobOwner != instAddr) {
		AltDB_DiagPushClient(slot, "HY010", "function sequence error");
		inst->status = dbERR_DATABASE; inst->dbError = DB_SQL_ERROR; return;
	}

	AltDB_GetData(slot, inst->columnIdx, inst->dataType, inst->pData, inst->dataSize,
	                &inst->status, &inst->dbError, &inst->actDataSize);
}
```

#### Disconnect.c - dbDisconnect
```c
/********************************************************************
 * Library: AltDB
 * File: Disconnect.c
 ********************************************************************
 * dbDisconnect (Section 7.10). Works regardless of connection state
 * (including BROKEN/FAILED) and takes the slot over from whichever
 * instance currently holds it, since tearing a connection down must
 * not be blockable by a stuck job on another instance.
 ********************************************************************/
#include <bur/plctypes.h>
#include <runtime.h>
#include <AsTCP.h>
#include <AltDB.h>
#include "Common.h"

void dbDisconnect(struct dbDisconnect *inst)
{
	UDINT instAddr = (UDINT)inst;
	UDINT slot;
	UINT generation;
	BOOL continuing;
	INT r;

	if (!inst->enable) {
		if (AltDB_SlotFromHandle(inst->connectionIdent, &slot, &generation) &&
		    gConn[slot].JobKind == JOB_DISCONNECT && gConn[slot].JobOwner == instAddr) {
			AltDB_Unlock(slot);
		}
		inst->status = ERR_FUB_ENABLE_FALSE; inst->dbError = 0;
		return;
	}

	if (!AltDB_SlotFromHandle(inst->connectionIdent, &slot, &generation)) {
		inst->status = dbERR_INVALID_HANDLE; inst->dbError = DB_SQL_INVALID_HANDLE; return;
	}

	continuing = gConn[slot].Locked && gConn[slot].JobKind == JOB_DISCONNECT && gConn[slot].JobOwner == instAddr;
	if (!continuing) {
		gConn[slot].Locked = TRUE;
		gConn[slot].JobOwner = instAddr;
		gConn[slot].JobKind = JOB_DISCONNECT;
	}

	r = AltDB_NetDisconnectStep(slot);
	if (r == NET_IN_PROGRESS) { inst->status = ERR_FUB_BUSY; return; }

	/* invalidate the handle (bump generation) before releasing the slot */
	gConn[slot].Generation = (UINT)((gConn[slot].Generation + 1) & 0x0FFF);
	AltDB_SlotReset(slot);

	inst->status = ERR_OK; inst->dbError = 0;
}
```

#### Info.c - dbGetInfo, dbGetErrorMessage
```c
/********************************************************************
 * Library: AltDB
 * File: Info.c
 ********************************************************************
 * dbGetInfo, dbGetErrorMessage (Section 7.11).
 *
 * dbGetInfo implements the small set of string info types that can
 * be answered from session data already held by the connection
 * (DBMS name/version, driver name/version, database name). All
 * other info types - including every numeric SQL_* capability flag
 * of Appendix A - are reported as dbERR_NOT_AVAILABLE, which Section
 * 7.11 documents as the correct response for an unsupported info
 * type, so this is a spec-compliant (if intentionally minimal)
 * implementation rather than a stub.
 ********************************************************************/
#include <bur/plctypes.h>
#include <runtime.h>
#include <AsTCP.h>
#include <AltDB.h>
#include "Common.h"
#include <string.h>

void dbGetInfo(struct dbGetInfo *inst)
{
	UDINT instAddr = (UDINT)inst;
	UDINT slot;
	UINT generation;
	const char *text;

	if (!inst->enable) { inst->status = ERR_FUB_ENABLE_FALSE; inst->dbError = 0; return; }
	if (!AltDB_SlotFromHandle(inst->connectionIdent, &slot, &generation)) {
		inst->status = dbERR_INVALID_HANDLE; inst->dbError = DB_SQL_INVALID_HANDLE; return;
	}
	if (gConn[slot].Locked && gConn[slot].JobOwner != instAddr) { inst->status = ERR_FUB_BUSY; return; }

	switch (inst->infoType) {
	case DB_IT_SQL_DBMS_NAME:    text = "Microsoft SQL Server"; break;
	case DB_IT_SQL_DBMS_VER:     text = gConn[slot].ServerVersion; break;
	case DB_IT_SQL_DRIVER_NAME:  text = "AltDB"; break;
	case DB_IT_SQL_DRIVER_VER:   text = "1.0.0000"; break;
	case DB_IT_SQL_DATABASE_NAME: text = gConn[slot].LoginDb; break;
	default: text = 0; break;
	}

	if (text == 0) {
		inst->status = dbERR_NOT_AVAILABLE; inst->dbError = DB_SQL_ERROR;
		return;
	}
	{
		UDINT n = (UDINT)strlen(text);
		UDINT need = n + 1;

		if (inst->serverInfoSize < need) {
			if (inst->pServerInfo != 0 && inst->serverInfoSize > 0) {
				UDINT copyLen = inst->serverInfoSize - 1;
				memcpy((void *)inst->pServerInfo, text, copyLen);
				((char *)inst->pServerInfo)[copyLen] = 0;
			}
			inst->status = dbERR_BUFFER_SIZE; inst->dbError = DB_SQL_ERROR;
			inst->actServerInfoSize = (UINT)need;
			return;
		}
		if (inst->pServerInfo != 0) memcpy((void *)inst->pServerInfo, text, need);
		inst->status = ERR_OK; inst->dbError = 0;
		inst->actServerInfoSize = (UINT)need;
	}
}

void dbGetErrorMessage(struct dbGetErrorMessage *inst)
{
	UDINT instAddr = (UDINT)inst;
	UDINT slot;
	UINT generation;
	DiagRec *rec;
	UDINT need;

	if (!inst->enable) { inst->status = ERR_FUB_ENABLE_FALSE; inst->dbError = 0; return; }
	if (!AltDB_SlotFromHandle(inst->connectionIdent, &slot, &generation)) {
		inst->status = dbERR_INVALID_HANDLE; inst->dbError = DB_SQL_INVALID_HANDLE; return;
	}
	/* available even while the connection is locked by another job or
	 * BROKEN/FAILED, mirroring AsDb's always-on diagnostics access */

	if (gConn[slot].DiagReadIdx >= gConn[slot].DiagCount) {
		memset(inst->sqlState, 0, sizeof(inst->sqlState));
		inst->nativeError = 0;
		inst->actErrorMessageSize = 0;
		inst->status = ERR_OK; inst->dbError = DB_SQL_NO_DATA;
		return;
	}

	rec = &gConn[slot].Diag[gConn[slot].DiagReadIdx];
	need = (UDINT)rec->MessageLen + 1;

	if (inst->errorMessageSize < need) {
		if (inst->pErrorMessage != 0 && inst->errorMessageSize > 0) {
			UDINT copyLen = inst->errorMessageSize - 1;
			memcpy((void *)inst->pErrorMessage, rec->Message, copyLen);
			((char *)inst->pErrorMessage)[copyLen] = 0;
		}
		memcpy(inst->sqlState, rec->SqlState, 6);
		inst->nativeError = rec->NativeError;
		inst->actErrorMessageSize = (INT)need;
		inst->status = dbERR_BUFFER_SIZE; inst->dbError = DB_SQL_ERROR;
		return; /* record remains unread, same contract as dbGetData */
	}

	if (inst->pErrorMessage != 0) memcpy((void *)inst->pErrorMessage, rec->Message, need);
	memcpy(inst->sqlState, rec->SqlState, 6);
	inst->nativeError = rec->NativeError;
	inst->actErrorMessageSize = (INT)need;
	inst->status = ERR_OK;
	inst->dbError = rec->IsError ? -1 : 1;
	gConn[slot].DiagReadIdx++;
}
```

#### ConnState.c - dbGetConnState (extension, diagnostic connection state snapshot)
```c
/********************************************************************
 * Library: AltDB
 * File: ConnState.c
 ********************************************************************
 * dbGetConnState (Section 7.12, extension FB - not part of AsDb).
 * Synchronous: returns a snapshot of the internal connection state
 * machine so a connection that appears stuck (e.g. a dbConnect/
 * dbExecuteSql/dbFetchNextRow call that keeps returning
 * ERR_FUB_BUSY) can be diagnosed from the calling IEC/C program
 * without instrumenting this library's C sources.
 ********************************************************************/
#include <bur/plctypes.h>
#include <runtime.h>
#include <AsTCP.h>
#include <AltDB.h>
#include "Common.h"
#include <string.h>

void dbGetConnState(struct dbGetConnState *inst)
{
	UDINT slot;
	UINT generation;
	ConnSlot *c;
	UDINT n;

	if (!inst->enable) { inst->status = ERR_FUB_ENABLE_FALSE; inst->dbError = 0; return; }
	if (!AltDB_SlotFromHandle(inst->connectionIdent, &slot, &generation)) {
		inst->status = dbERR_INVALID_HANDLE; inst->dbError = DB_SQL_INVALID_HANDLE; return;
	}

	c = &gConn[slot];
	memset(&inst->connState, 0, sizeof(inst->connState));

	inst->connState.state = c->State;
	inst->connState.netStep = c->NetStep;
	inst->connState.jobKind = c->JobKind;
	inst->connState.locked = c->Locked;
	inst->connState.tcpIdent = c->TcpIdent;
	inst->connState.encoding = c->Encoding;
	inst->connState.packetSize = c->PacketSize;
	inst->connState.sendLen = c->SendLen;
	inst->connState.sendPos = c->SendPos;
	inst->connState.tokLen = c->TokLen;
	inst->connState.tokPos = c->TokPos;
	inst->connState.statementActive = c->StatementActive;
	inst->connState.columnCount = c->ColumnCount;
	inst->connState.hasResultSet = c->HasResultSet;
	inst->connState.resultSetOpen = c->ResultSetOpen;
	inst->connState.rowReady = c->RowReady;
	inst->connState.noMoreRows = c->NoMoreRows;
	inst->connState.affectedRows = c->AffectedRows;
	inst->connState.affectedRowsKnown = c->AffectedRowsKnown;
	inst->connState.diagCount = c->DiagCount;
	inst->connState.diagReadIdx = c->DiagReadIdx;

	/* IEC STRING[31] is generated as a plain NUL-terminated char[32]
	 * (confirmed against AsTCP.h's AsTcpMcsType.name), not a
	 * length-prefixed Pascal string. */
	n = (UDINT)strlen(c->ServerVersion);
	if (n > 31) n = 31;
	memcpy((char *)&inst->connState.serverVersion, c->ServerVersion, n);
	((char *)&inst->connState.serverVersion)[n] = 0;

	inst->status = ERR_OK;
	inst->dbError = 0;
}
```

### Program Logical/AltDBExample (IEC)

#### Main.st - Init, cyclic, exit code
```iecst
(********************************************************************
 * COPYRIGHT --
 ********************************************************************
 * Program: SQLRecipe
 * File: SQLRecipe.st
 * Author: B&R
 * Created: December 27, 2010
 ********************************************************************
 * Implementation of program SQLRecipe
 ********************************************************************)

PROGRAM _INIT

(* TODO : Add your code here *)

END_PROGRAM

PROGRAM _CYCLIC

	CASE Command.eCommand OF
		eCMD_IDLE :
		eCMD_CONNECT :
			IF eStep = eSTOP THEN
				eStep := eCONNECT;
				Command.eCommand := eCMD_CONNECT_w;
			END_IF
		eCMD_CONNECT_w:
			IF eStep = eWAIT_FOR_COMMAND THEN
				Command.eCommand := eCMD_IDLE;
			END_IF
		eCMD_LOAD :
			IF eStep = eWAIT_FOR_COMMAND THEN
				eStep := eLOAD_RECEIPE;
				Command.eCommand := eCMD_LOAD_w;
			END_IF
		eCMD_LOAD_w:
			IF eStep = eWAIT_FOR_COMMAND THEN
				Command.eCommand := eCMD_IDLE;
			END_IF
		eCMD_SAVE :
			IF eStep = eWAIT_FOR_COMMAND THEN
				eStep := eSAVE_RECEIPE;
				Command.eCommand := eCMD_SAVE_w;
			END_IF
		eCMD_SAVE_w:
			IF eStep = eWAIT_FOR_COMMAND THEN
				Command.eCommand := eCMD_IDLE;
			END_IF
		eCMD_SAVEAS :
			IF eStep = eWAIT_FOR_COMMAND THEN
				eStep := eSAVE_AS;
				Command.eCommand := eCMD_SAVEAS_w;
			END_IF
		eCMD_SAVEAS_w:
			IF eStep = eWAIT_FOR_COMMAND THEN
				Command.eCommand := eCMD_IDLE;
			END_IF
		eCMD_DELETE :
			IF eStep = eWAIT_FOR_COMMAND THEN
				eStep := eDELETE_RECEIPE;
				Command.eCommand := eCMD_DELETE_w;
			END_IF
		eCMD_DELETE_w:
			IF eStep = eWAIT_FOR_COMMAND THEN
				Command.eCommand := eCMD_IDLE;
			END_IF
		eCMD_RENAME :
			IF eStep = eWAIT_FOR_COMMAND THEN
				eStep := eRENAME_RECEIPE;
				Command.eCommand := eCMD_RENAME_w;
			END_IF
		eCMD_RENAME_w:
			IF eStep = eWAIT_FOR_COMMAND THEN
				Command.eCommand := eCMD_IDLE;
			END_IF
		eCMD_DISCONNECT :
			IF eStep = eWAIT_FOR_COMMAND OR
				eStep = eERROR THEN
				eStep := eDISCONNECT;
				Command.eCommand := eCMD_DISCONNECT_w;
			END_IF
		eCMD_DISCONNECT_w:
			IF eStep = eSTOP THEN
				Command.eCommand := eCMD_IDLE;
			END_IF
	END_CASE

	CASE eStep OF
		(* connect to database *)
		eCONNECT :
			brsmemset( ADR(ReceipeDBConnect), 0, SIZEOF(ReceipeDBConnect) );
			ReceipeDBConnect.enable := TRUE;
			ReceipeDBConnect.databaseSystem := DB_SYSTEM_MS_SQL;
			ReceipeDBConnect.pUserName := ADR(USERNAME);
			ReceipeDBConnect.pPassword := ADR(PASSWORD);
			ReceipeDBConnect.pServerName := ADR(HOST);
			ReceipeDBConnect.pDatabaseName := ADR(DATABASE);
			eStep := eCONNECT_r;
		eCONNECT_r :
			ReceipeDBConnect();
			IF ReceipeDBConnect.status = 0 THEN
				ConnectionIdent := ReceipeDBConnect.connectionIdent;
				eStep := eGET_TABLES;
			ELSIF ReceipeDBConnect.status <> 65535 THEN
				IF ReceipeDBConnect.connectionIdent <> 0 THEN
					ConnectionIdent := ReceipeDBConnect.connectionIdent;
					eStep := eGET_ERROR;
				ELSE
					eStep := eERROR;
				END_IF
			END_IF

			(* read out available tables *)
		eGET_TABLES :
			brsstrcpy( ADR(sSQLstring), ADR('SELECT name FROM sysobjects WHERE type=$'u$'') );
			ReceipeDBExecute.enable := TRUE;
			ReceipeDBExecute.pSqlStatement := ADR(sSQLstring);
			ReceipeDBExecute.connectionIdent := ConnectionIdent;
			eStep := eGET_TABLES_r;
		eGET_TABLES_r :
			ReceipeDBExecute();
			IF ReceipeDBExecute.status = ERR_OK THEN
				eStep := eFETCH_NEXT_ROW;
			ELSIF ReceipeDBExecute.status <> ERR_FUB_BUSY THEN
				eStep := eGET_ERROR;
			END_IF
			(* prepare one row to read column(s) *)
		eFETCH_NEXT_ROW :
			ReceipeDBFetchNextRow.enable := TRUE;
			ReceipeDBFetchNextRow.connectionIdent := ConnectionIdent;
			eStep := eFETCH_NEXT_ROW_r;
		eFETCH_NEXT_ROW_r :
			ReceipeDBFetchNextRow();
			IF ReceipeDBFetchNextRow.status = ERR_OK THEN
				eStep := eREAD_TABLE_NAME;
			ELSIF ReceipeDBFetchNextRow.status <> ERR_FUB_BUSY THEN
				IF ReceipeDBFetchNextRow.dbError = 100 THEN
					eStep := eCREATE_TABLE;
				ELSE
					eStep := eGET_ERROR;
				END_IF
			END_IF
			(* read out 1st column -> name *)
		eREAD_TABLE_NAME :
			ReceipeDBGetData.enable := TRUE;
			ReceipeDBGetData.connectionIdent := ConnectionIdent;
			ReceipeDBGetData.columnIdx := 1;
			ReceipeDBGetData.pData := ADR( sData );
			ReceipeDBGetData.dataSize := SIZEOF( sData );
			ReceipeDBGetData.dataType := DB_SQL_CHAR;
			eStep := eREAD_TABLE_NAME_r;
		eREAD_TABLE_NAME_r :
			ReceipeDBGetData();
			IF ReceipeDBGetData.status = 0 THEN
				IF brsstrcmp( ADR(sData), ADR(TABLE) )=0 THEN
					eStep := eGET_RECEIPE_NAMES;
				ELSE
					eStep := eFETCH_NEXT_ROW;
				END_IF
			ELSIF ReceipeDBGetData.status <> ERR_FUB_BUSY THEN
				eStep := eGET_ERROR;
			END_IF

			(* Create New Table *)
		eCREATE_TABLE :
			brsstrcpy( ADR(sSQLstring), ADR('CREATE TABLE '));
			brsstrcat( ADR(sSQLstring), ADR(TABLE));
			brsstrcat( ADR(sSQLstring), ADR(' (') );
			brsstrcat( ADR(sSQLstring), ADR('idx smallint IDENTITY (1,1) PRIMARY KEY, ') );
			brsstrcat( ADR(sSQLstring), ADR('name varchar(') );
			brsitoa(LENGTH_NAME, ADR(sSQLstring) + brsstrlen(ADR(sSQLstring)) );
			brsstrcat( ADR(sSQLstring), ADR(') UNIQUE, ') );
			brsstrcat( ADR(sSQLstring), ADR('price real, ') );
			brsstrcat( ADR(sSQLstring), ADR('setTemp real, ') );
			brsstrcat( ADR(sSQLstring), ADR('milk real, ') );
			brsstrcat( ADR(sSQLstring), ADR('sugar real, ') );
			brsstrcat( ADR(sSQLstring), ADR('coffee real, ') );
			brsstrcat( ADR(sSQLstring), ADR('water real ') );
			brsstrcat( ADR(sSQLstring), ADR(')') );
			ReceipeDBExecute.enable := TRUE;
			ReceipeDBExecute.pSqlStatement := ADR(sSQLstring);
			ReceipeDBExecute.connectionIdent := ConnectionIdent;
			eStep := eCREATE_TABLE_r;
		eCREATE_TABLE_r :
			ReceipeDBExecute();
			IF ReceipeDBExecute.status = ERR_OK THEN
				eStep := eINSERT_DEFAULT;
			ELSIF ReceipeDBExecute.status <> ERR_FUB_BUSY THEN
				eStep := eGET_ERROR;
			END_IF
			(* fill default receipe *)
		eINSERT_DEFAULT :
			brsstrcpy( ADR(sSQLstring), ADR('INSERT INTO ') );
			brsstrcat( ADR(sSQLstring), ADR(TABLE) );
			brsstrcat( ADR(sSQLstring), ADR(' (name, price, setTemp, milk, sugar, coffee, water) ') );
			brsstrcat( ADR(sSQLstring), ADR(' VALUES ($'default$',$'1.73$',$'80.0$',$'95.0$',$'33.3$',$'66.6$',$'155.3$')') );
			ReceipeDBExecute.enable := TRUE;
			ReceipeDBExecute.pSqlStatement := ADR(sSQLstring);
			ReceipeDBExecute.connectionIdent := ConnectionIdent;
			eStep := eINSERT_DEFAULT_r;
		eINSERT_DEFAULT_r :
			ReceipeDBExecute();
			IF ReceipeDBExecute.status = ERR_OK THEN
				eStep := eGET_RECEIPE_NAMES;
			ELSIF ReceipeDBExecute.status <> ERR_FUB_BUSY THEN
				eStep := eGET_ERROR;
			END_IF

			(* get receipe names - only as much as can saved in list *)
		eGET_RECEIPE_NAMES :
			brsstrcpy( ADR(sSQLstring), ADR('SELECT TOP(') );
			brsitoa( SIZEOF(Command.sReceipeNames)/SIZEOF(Command.sReceipeNames[0]), ADR(sSQLstring) + brsstrlen(ADR(sSQLstring)) );
			brsstrcat( ADR(sSQLstring), ADR(') name FROM ') );
			brsstrcat( ADR(sSQLstring), ADR(TABLE) );
			brsstrcat( ADR(sSQLstring), ADR(' ORDER BY name ASC') );
			ReceipeDBExecute.enable := TRUE;
			ReceipeDBExecute.pSqlStatement := ADR(sSQLstring);
			ReceipeDBExecute.connectionIdent := ConnectionIdent;
			ReceipeNameCounter := 0;
			brsmemset( ADR(Command.sReceipeNames), 0, SIZEOF(Command.sReceipeNames) );
			eStep := eGET_RECEIPE_NAMES_r;
		eGET_RECEIPE_NAMES_r:
			ReceipeDBExecute();
			IF ReceipeDBExecute.status = ERR_OK THEN
				eStep := eFETCH_RECEIPE_NAME;
			ELSIF ReceipeDBExecute.status <> ERR_FUB_BUSY THEN
				eStep := eGET_ERROR;
			END_IF
			(* prepare one row to read column(s) *)
		eFETCH_RECEIPE_NAME :
			ReceipeDBFetchNextRow.enable := TRUE;
			ReceipeDBFetchNextRow.connectionIdent := ConnectionIdent;
			eStep := eFETCH_RECEIPE_NAME_r;
		eFETCH_RECEIPE_NAME_r :
			ReceipeDBFetchNextRow();
			IF ReceipeDBFetchNextRow.status = ERR_OK THEN
				eStep := eREAD_RECEIPE_NAME;
			ELSIF ReceipeDBFetchNextRow.status <> ERR_FUB_BUSY THEN
				IF ReceipeDBFetchNextRow.dbError = DB_SQL_NO_DATA THEN
					IF ReceipeNameCounter = 0 THEN	(* no receipe - maybe last receipe deleted *)
						eStep := eINSERT_DEFAULT;
					ELSE
						eStep := eWAIT_FOR_COMMAND;	(* all receipes read - wait for command *)
					END_IF
				ELSE
					eStep := eGET_ERROR;
				END_IF
			END_IF
			(* read out 1st column -> name *)
		eREAD_RECEIPE_NAME :
			ReceipeDBGetData.enable := TRUE;
			ReceipeDBGetData.connectionIdent := ConnectionIdent;
			ReceipeDBGetData.columnIdx := 1;
			ReceipeDBGetData.pData := ADR( Command.sReceipeNames[ReceipeNameCounter] );
			ReceipeDBGetData.dataSize := SIZEOF(Command.sReceipeNames[0]) - 1;
			ReceipeDBGetData.dataType := DB_SQL_CHAR;
			eStep := eREAD_RECEIPE_NAME_r;
		eREAD_RECEIPE_NAME_r :
			ReceipeDBGetData();
			IF ReceipeDBGetData.status = 0 THEN
				ReceipeNameCounter := ReceipeNameCounter + 1;
				IF ReceipeNameCounter < (SIZEOF(Command.sReceipeNames)/SIZEOF(Command.sReceipeNames[0])) THEN
					eStep := eFETCH_RECEIPE_NAME;
				ELSE
					Command.uStatus := 0;
					eStep := eWAIT_FOR_COMMAND;
				END_IF
			ELSIF ReceipeDBGetData.status <> ERR_FUB_BUSY THEN
				eStep := eGET_ERROR;
			END_IF

		eWAIT_FOR_COMMAND :

			(* Load a receipe *)
		eLOAD_RECEIPE :
			brsstrcpy( ADR(sSQLstring), ADR('SELECT price, setTemp, milk, sugar, coffee, water FROM ') );
			brsstrcat( ADR(sSQLstring), ADR(TABLE) );
			brsstrcat( ADR(sSQLstring), ADR(' WHERE name = $'') );
			brsstrcat( ADR(sSQLstring), ADR(Command.sNewReceipe) );
			brsstrcat( ADR(sSQLstring), ADR('$'') );
			ReceipeDBExecute.enable := TRUE;
			ReceipeDBExecute.pSqlStatement := ADR(sSQLstring);
			ReceipeDBExecute.connectionIdent := ConnectionIdent;
			eStep := eLOAD_RECEIPE_r;
		eLOAD_RECEIPE_r :
			ReceipeDBExecute();
			IF ReceipeDBExecute.status = ERR_OK THEN
				eStep := eFETCH_VALUES;
			ELSIF ReceipeDBExecute.status <> ERR_FUB_BUSY THEN
				IF ReceipeDBExecute.dbError = 100 THEN
					eStep := eWAIT_FOR_COMMAND;
				ELSE
					eStep := eGET_ERROR;
				END_IF
			END_IF
			(* prepare one row to read column(s) *)
		eFETCH_VALUES :
			ReceipeDBFetchNextRow.enable := TRUE;
			ReceipeDBFetchNextRow.connectionIdent := ConnectionIdent;
			eStep := eFETCH_VALUES_r;
		eFETCH_VALUES_r :
			ReceipeDBFetchNextRow();
			IF ReceipeDBFetchNextRow.status = ERR_OK THEN
				usCol := 1;
				eStep := eGET_VALUES;
			ELSIF ReceipeDBFetchNextRow.status <> ERR_FUB_BUSY THEN
				IF ReceipeDBFetchNextRow.dbError = DB_SQL_NO_DATA THEN
					Command.uStatus := 1;
					eStep := eWAIT_FOR_COMMAND;
				ELSE
					eStep := eGET_ERROR;
				END_IF
			END_IF
			(* read out all columns *)
		eGET_VALUES :
			ReceipeDBGetData.enable := TRUE;
			ReceipeDBGetData.connectionIdent := ConnectionIdent;
			ReceipeDBGetData.columnIdx := usCol;
			CASE usCol OF
				1:
					ReceipeDBGetData.pData := ADR(gMainLogic.par.receipe.price);
					ReceipeDBGetData.dataSize := SIZEOF(gMainLogic.par.receipe.price);
					ReceipeDBGetData.dataType := DB_SQL_REAL;
				2:
					ReceipeDBGetData.pData := ADR(gMainLogic.par.receipe.setTemp);
					ReceipeDBGetData.dataSize := SIZEOF(gMainLogic.par.receipe.setTemp);
					ReceipeDBGetData.dataType := DB_SQL_REAL;
				3:
					ReceipeDBGetData.pData := ADR(gMainLogic.par.receipe.milk);
					ReceipeDBGetData.dataSize := SIZEOF(gMainLogic.par.receipe.milk);
					ReceipeDBGetData.dataType := DB_SQL_REAL;
				4:
					ReceipeDBGetData.pData := ADR(gMainLogic.par.receipe.sugar);
					ReceipeDBGetData.dataSize := SIZEOF(gMainLogic.par.receipe.sugar);
					ReceipeDBGetData.dataType := DB_SQL_REAL;
				5:
					ReceipeDBGetData.pData := ADR(gMainLogic.par.receipe.coffee);
					ReceipeDBGetData.dataSize := SIZEOF(gMainLogic.par.receipe.coffee);
					ReceipeDBGetData.dataType := DB_SQL_REAL;
				6:
					ReceipeDBGetData.pData := ADR(gMainLogic.par.receipe.water);
					ReceipeDBGetData.dataSize := SIZEOF(gMainLogic.par.receipe.water);
					ReceipeDBGetData.dataType := DB_SQL_REAL;
			END_CASE
			eStep := eGET_VALUES_r;
		eGET_VALUES_r :
			ReceipeDBGetData();
			IF ReceipeDBGetData.status = 0 THEN
				usCol := usCol + 1;
				IF usCol <= 6 THEN
					eStep := eGET_VALUES;
				ELSE
					Command.uStatus := ERR_OK;
					brsstrcpy( ADR(Command.sActReceipe), ADR(Command.sNewReceipe) );
					eStep := eWAIT_FOR_COMMAND;
				END_IF
			ELSIF ReceipeDBGetData.status <> ERR_FUB_BUSY THEN
				eStep := eGET_ERROR;
			END_IF

			(* save receipe *)
		eSAVE_RECEIPE :
			brsstrcpy( ADR(sSQLstring), ADR('UPDATE ') );
			brsstrcat( ADR(sSQLstring), ADR(TABLE) );
			brsstrcat( ADR(sSQLstring), ADR(' SET price=$'') );
			brsftoa( gMainLogic.par.receipe.price, ADR(sSQLstring) + brsstrlen(ADR(sSQLstring)) );
			brsstrcat( ADR(sSQLstring), ADR('$', setTemp=$'') );
			brsftoa( gMainLogic.par.receipe.setTemp, ADR(sSQLstring) + brsstrlen(ADR(sSQLstring)) );
			brsstrcat( ADR(sSQLstring), ADR('$', milk=$'') );
			brsftoa( gMainLogic.par.receipe.milk, ADR(sSQLstring) + brsstrlen(ADR(sSQLstring)) );
			brsstrcat( ADR(sSQLstring), ADR('$', sugar=$'') );
			brsftoa( gMainLogic.par.receipe.sugar, ADR(sSQLstring) + brsstrlen(ADR(sSQLstring)) );
			brsstrcat( ADR(sSQLstring), ADR('$', coffee=$'') );
			brsftoa( gMainLogic.par.receipe.coffee, ADR(sSQLstring) + brsstrlen(ADR(sSQLstring)) );
			brsstrcat( ADR(sSQLstring), ADR('$', water=$'') );
			brsftoa( gMainLogic.par.receipe.water, ADR(sSQLstring) + brsstrlen(ADR(sSQLstring)) );
			brsstrcat( ADR(sSQLstring), ADR('$' WHERE name=$'') );
			brsstrcat( ADR(sSQLstring), ADR(Command.sActReceipe) );
			brsstrcat( ADR(sSQLstring), ADR('$'') );
			ReceipeDBExecute.enable := TRUE;
			ReceipeDBExecute.pSqlStatement := ADR(sSQLstring);
			ReceipeDBExecute.connectionIdent := ConnectionIdent;
			eStep := eSAVE_RECEIPE_r;
		eSAVE_RECEIPE_r :
			ReceipeDBExecute();
			IF ReceipeDBExecute.status = ERR_OK THEN
				eStep := eSAVE_GET_AFFECTED_ROWS;
			ELSIF ReceipeDBExecute.status <> ERR_FUB_BUSY THEN
				eStep := eGET_ERROR;
			END_IF
			(* test if on row is saved *)
		eSAVE_GET_AFFECTED_ROWS :
			ReceipeDBGetAffectedRows.enable := TRUE;
			ReceipeDBGetAffectedRows.connectionIdent := ConnectionIdent;
			eStep := eSAVE_GET_AFFECTED_ROWS_r;
		eSAVE_GET_AFFECTED_ROWS_r :
			ReceipeDBGetAffectedRows();
			IF ReceipeDBGetAffectedRows.status = ERR_OK THEN
				IF ReceipeDBGetAffectedRows.affectedRows = 1 THEN	(* one row updated -> correct *)
					Command.uStatus := 0;
				ELSE
					Command.uStatus := 1;
				END_IF
				eStep := eWAIT_FOR_COMMAND;
			ELSIF ReceipeDBGetAffectedRows.status <> ERR_FUB_BUSY THEN
				eStep := eGET_ERROR;
			END_IF

			(* save with new name *)
			(* only if not exist *)
		eSAVE_AS :
			brsstrcpy( ADR(sSQLstring), ADR('IF NOT EXISTS (SELECT * FROM ') );
			brsstrcat( ADR(sSQLstring), ADR(TABLE) );
			brsstrcat( ADR(sSQLstring), ADR(' WHERE name=$'') );
			brsstrcat( ADR(sSQLstring), ADR(Command.sNewReceipe) );
			brsstrcat( ADR(sSQLstring), ADR('$') ') );
			brsstrcat( ADR(sSQLstring), ADR('INSERT INTO ') );
			brsstrcat( ADR(sSQLstring), ADR(TABLE) );
			brsstrcat( ADR(sSQLstring), ADR(' (name, price, setTemp, milk, sugar, coffee, water) ') );
			brsstrcat( ADR(sSQLstring), ADR('VALUES ($'') );
			brsstrcat( ADR(sSQLstring), ADR(Command.sNewReceipe) );
			brsstrcat( ADR(sSQLstring), ADR('$',$'') );
			brsftoa( gMainLogic.par.receipe.price, ADR(sSQLstring) + brsstrlen(ADR(sSQLstring)) );
			brsstrcat( ADR(sSQLstring), ADR('$',$'') );
			brsftoa( gMainLogic.par.receipe.setTemp, ADR(sSQLstring) + brsstrlen(ADR(sSQLstring)) );
			brsstrcat( ADR(sSQLstring), ADR('$',$'') );
			brsftoa( gMainLogic.par.receipe.milk, ADR(sSQLstring) + brsstrlen(ADR(sSQLstring)) );
			brsstrcat( ADR(sSQLstring), ADR('$',$'') );
			brsftoa( gMainLogic.par.receipe.sugar, ADR(sSQLstring) + brsstrlen(ADR(sSQLstring)) );
			brsstrcat( ADR(sSQLstring), ADR('$',$'') );
			brsftoa( gMainLogic.par.receipe.coffee, ADR(sSQLstring) + brsstrlen(ADR(sSQLstring)) );
			brsstrcat( ADR(sSQLstring), ADR('$',$'') );
			brsftoa( gMainLogic.par.receipe.water, ADR(sSQLstring) + brsstrlen(ADR(sSQLstring)) );
			brsstrcat( ADR(sSQLstring), ADR('$')') );
			ReceipeDBExecute.enable := TRUE;
			ReceipeDBExecute.pSqlStatement := ADR(sSQLstring);
			ReceipeDBExecute.connectionIdent := ConnectionIdent;
			eStep := eSAVE_AS_r;
		eSAVE_AS_r :
			ReceipeDBExecute();
			IF ReceipeDBExecute.status = ERR_OK THEN
				eStep := eSAVE_AS_ROWS_AFFECTED;
			ELSIF ReceipeDBExecute.status <> ERR_FUB_BUSY THEN
				eStep := eGET_ERROR;
			END_IF
			(* test if on row is changed *)
		eSAVE_AS_ROWS_AFFECTED :
			ReceipeDBGetAffectedRows.enable := TRUE;
			ReceipeDBGetAffectedRows.connectionIdent := ConnectionIdent;
			eStep := eSAVE_AS_ROWS_AFFECTED_r;
		eSAVE_AS_ROWS_AFFECTED_r :
			ReceipeDBGetAffectedRows();
			IF ReceipeDBGetAffectedRows.status = ERR_OK THEN
				IF ReceipeDBGetAffectedRows.affectedRows = 1 THEN	(* one row updated -> correct *)
					Command.uStatus := 0;
					brsstrcpy( ADR(Command.sActReceipe), ADR(Command.sNewReceipe) );
				ELSE
					Command.uStatus := 1;
					brsstrcpy( ADR(Command.sActReceipe), ADR('') );
				END_IF
				eStep := eGET_RECEIPE_NAMES;
			ELSIF ReceipeDBGetAffectedRows.status <> ERR_FUB_BUSY THEN
				eStep := eGET_ERROR;
			END_IF

			(* delete receipe *)
		eDELETE_RECEIPE :
			brsstrcpy( ADR(sSQLstring), ADR('DELETE FROM ') );
			brsstrcat( ADR(sSQLstring), ADR(TABLE) );
			brsstrcat( ADR(sSQLstring), ADR(' WHERE name=$'') );
			brsstrcat( ADR(sSQLstring), ADR(Command.sNewReceipe) );
			brsstrcat( ADR(sSQLstring), ADR('$'') );
			ReceipeDBExecute.enable := TRUE;
			ReceipeDBExecute.pSqlStatement := ADR(sSQLstring);
			ReceipeDBExecute.connectionIdent := ConnectionIdent;
			eStep := eDELETE_RECEIPE_r;
		eDELETE_RECEIPE_r :
			ReceipeDBExecute();
			IF ReceipeDBExecute.status = ERR_OK THEN
				eStep := eDELETE_ROWS_AFFECTED;
			ELSIF ReceipeDBExecute.status <> ERR_FUB_BUSY THEN
				eStep := eGET_ERROR;
			END_IF
			(* test if on row is changed *)
		eDELETE_ROWS_AFFECTED :
			ReceipeDBGetAffectedRows.enable := TRUE;
			ReceipeDBGetAffectedRows.connectionIdent := ConnectionIdent;
			eStep := eDELETE_ROWS_AFFECTED_r;
		eDELETE_ROWS_AFFECTED_r :
			ReceipeDBGetAffectedRows();
			IF ReceipeDBGetAffectedRows.status = ERR_OK THEN
				IF ReceipeDBGetAffectedRows.affectedRows = 1 THEN	(* one row updated -> correct *)
					Command.uStatus := 0;
					IF brsstrcmp( ADR(Command.sActReceipe), ADR(Command.sNewReceipe) ) = 0 THEN	(* when delete actual receipe *)
						brsstrcpy( ADR(Command.sActReceipe), ADR('') );
					END_IF
					brsstrcpy( ADR(Command.sNewReceipe), ADR('') );
				ELSE
					Command.uStatus := 1;
				END_IF
				eStep := eGET_RECEIPE_NAMES;
			ELSIF ReceipeDBGetAffectedRows.status <> ERR_FUB_BUSY THEN
				eStep := eGET_ERROR;
			END_IF

			(* rename receipe *)
			(* only if new name not exist *)
		eRENAME_RECEIPE :
			brsstrcpy( ADR(sSQLstring), ADR('IF NOT EXISTS (SELECT * FROM ') );
			brsstrcat( ADR(sSQLstring), ADR(TABLE) );
			brsstrcat( ADR(sSQLstring), ADR(' WHERE name=$'') );
			brsstrcat( ADR(sSQLstring), ADR(Command.sNewReceipe) );
			brsstrcat( ADR(sSQLstring), ADR('$') ') );
			brsstrcat( ADR(sSQLstring), ADR('UPDATE ') );
			brsstrcat( ADR(sSQLstring), ADR(TABLE) );
			brsstrcat( ADR(sSQLstring), ADR(' SET name=$'') );
			brsstrcat( ADR(sSQLstring), ADR(Command.sNewReceipe) );
			brsstrcat( ADR(sSQLstring), ADR('$' WHERE name=$'') );
			brsstrcat( ADR(sSQLstring), ADR(Command.sActReceipe) );
			brsstrcat( ADR(sSQLstring), ADR('$'') );
			ReceipeDBExecute.enable := TRUE;
			ReceipeDBExecute.pSqlStatement := ADR(sSQLstring);
			ReceipeDBExecute.connectionIdent := ConnectionIdent;
			eStep := eRENAME_RECEIPE_r;
		eRENAME_RECEIPE_r :
			ReceipeDBExecute();
			IF ReceipeDBExecute.status = ERR_OK THEN
				eStep := eRENAME_GET_AFFECTED_ROWS;
			ELSIF ReceipeDBExecute.status <> ERR_FUB_BUSY THEN
				eStep := eGET_ERROR;
			END_IF
			(* test if on row is changed *)
		eRENAME_GET_AFFECTED_ROWS :
			ReceipeDBGetAffectedRows.enable := TRUE;
			ReceipeDBGetAffectedRows.connectionIdent := ConnectionIdent;
			eStep := eRENAME_GET_AFFECTED_ROWS_r;
		eRENAME_GET_AFFECTED_ROWS_r :
			ReceipeDBGetAffectedRows();
			IF ReceipeDBGetAffectedRows.status = ERR_OK THEN
				IF ReceipeDBGetAffectedRows.affectedRows = 1 THEN	(* one row updated -> correct *)
					Command.uStatus := 0;
					brsstrcpy( ADR(Command.sActReceipe),ADR(Command.sNewReceipe) );
				ELSE
					Command.uStatus := 1;
					brsstrcpy( ADR(Command.sActReceipe),ADR('') );
				END_IF
				eStep := eGET_RECEIPE_NAMES;
			ELSIF ReceipeDBGetAffectedRows.status <> ERR_FUB_BUSY THEN
				eStep := eGET_ERROR;
			END_IF

			(* disconnect from server *)
		eDISCONNECT :
			ReceipeDBDisconnect.enable := TRUE;
			ReceipeDBDisconnect.connectionIdent := ConnectionIdent;
			eStep := eDISCONNECT_r;
		eDISCONNECT_r :
			ReceipeDBDisconnect();
			IF ReceipeDBDisconnect.status <> ERR_FUB_BUSY THEN
				eStep := eSTOP;
				ConnectionIdent := 0;
			END_IF

			(* get error string *)
		eGET_ERROR :
			brsmemset( ADR(Command.sErrorString), 0, SIZEOF(Command.sErrorString) );
			ReceipeDBErrMsg.enable := TRUE;
			ReceipeDBErrMsg.connectionIdent := ConnectionIdent;
			ReceipeDBErrMsg.pErrorMessage := ADR( Command.sErrorString );
			ReceipeDBErrMsg.errorMessageSize := SIZEOF( Command.sErrorString ) - 1;
			eStep := eGET_ERROR_r;
		eGET_ERROR_r :
			ReceipeDBErrMsg();

			IF ReceipeDBErrMsg.status <> ERR_FUB_BUSY THEN
				Command.uStatus := 2;
				eStep := eERROR;
			END_IF
	END_CASE;
	DBConnectState();

END_PROGRAM

(********************************************************************
 * COPYRIGHT --
 ********************************************************************
 * Program: SQLRecipe
 * File: SQLRecipe_exit.st
 * Author: B&R
 * Created: January 04, 2011
 *******************************************************************)

PROGRAM _EXIT
	WHILE eStep <> eSTOP DO
		CASE eStep OF
			(* Finish dbConnect FUB befor close connection *)
			eCONNECT_r:
				ReceipeDBConnect();
				IF ReceipeDBConnect.status <> ERR_FUB_BUSY THEN
					eStep := eDISCONNECT;
				END_IF
				(* Finish dbExecuteSQL FUB *)
				eGET_TABLES_r,
				eCREATE_TABLE_r,
				eINSERT_DEFAULT_r,
				eGET_RECEIPE_NAMES_r,
				eLOAD_RECEIPE_r,
				eSAVE_RECEIPE_r,
				eSAVE_AS_r,
				eDELETE_RECEIPE_r,
			eRENAME_RECEIPE_r:
				ReceipeDBExecute();
				IF ReceipeDBExecute.status <> ERR_FUB_BUSY THEN
					eStep := eDISCONNECT;
				END_IF
				(* Finish dbGetAffectedRows FUB *)
				eSAVE_GET_AFFECTED_ROWS_r,
				eSAVE_AS_ROWS_AFFECTED_r,
				eDELETE_ROWS_AFFECTED_r,
			eRENAME_GET_AFFECTED_ROWS_r:
				ReceipeDBGetAffectedRows();
				IF ReceipeDBGetAffectedRows.status <> ERR_FUB_BUSY THEN
					eStep := eDISCONNECT;
				END_IF
				(* Finish dbFetchNextRow FUB *)
				eFETCH_NEXT_ROW_r,
				eFETCH_RECEIPE_NAME_r,
			eFETCH_VALUES_r:
				ReceipeDBFetchNextRow();
				IF ReceipeDBFetchNextRow.status <> ERR_FUB_BUSY THEN
					eStep := eDISCONNECT;
				END_IF
				(* Finish dbGetData FUB *)
				eREAD_TABLE_NAME_r,
				eREAD_RECEIPE_NAME_r,
			eGET_VALUES_r:
				ReceipeDBGetData();
				IF ReceipeDBGetData.status <> ERR_FUB_BUSY THEN
					eStep := eDISCONNECT;
				END_IF
				(* Finish dbGetErrorMessage FUB *)
			eGET_ERROR_r:
				ReceipeDBErrMsg();
				IF ReceipeDBErrMsg.status <> ERR_FUB_BUSY THEN
					eStep := eDISCONNECT;
				END_IF
				(* Disconnect *)
			eDISCONNECT:
				ReceipeDBDisconnect.enable := TRUE;
				ReceipeDBDisconnect.connectionIdent := ConnectionIdent;
				eStep := eDISCONNECT_r;
				(* Run Disconnect FUB *)
			eDISCONNECT_r:
				ReceipeDBDisconnect();
				IF ReceipeDBDisconnect.status <> ERR_FUB_BUSY THEN
					eStep := eSTOP;
				END_IF

			eERROR:
				eStep := eDISCONNECT;
			ELSE
				eStep := eDISCONNECT;
		END_CASE
	END_WHILE;
END_PROGRAM
```

#### Types.typ - Local data types
```iecst
(********************************************************************
 * COPYRIGHT --
 ********************************************************************
 * Program: SQLRecipe
 * File: SQLRecipe.typ
 * Author: B&R
 * Created: December 27, 2010
 ********************************************************************
 * Local data types of program SQLRecipe
 ********************************************************************)

TYPE
	Steps_enum :
		(
		eSTOP, (*Stop - nothing to do*)
		eCONNECT, (*Connect to Database*)
		eCONNECT_r,
		eGET_TABLES, (*SELECT Names of Tables in Database*)
		eGET_TABLES_r,
		eFETCH_NEXT_ROW, (*Read line by line*)
		eFETCH_NEXT_ROW_r,
		eREAD_TABLE_NAME, (*Get name out of line*)
		eREAD_TABLE_NAME_r,
		eCREATE_TABLE, (*CREATE TABLE with name if not exist*)
		eCREATE_TABLE_r,
		eINSERT_DEFAULT, (*INSERT default receipe*)
		eINSERT_DEFAULT_r,
		eGET_RECEIPE_NAMES := 30, (*SELECT Names of all receipes*)
		eGET_RECEIPE_NAMES_r,
		eFETCH_RECEIPE_NAME, (*read line by line*)
		eFETCH_RECEIPE_NAME_r,
		eREAD_RECEIPE_NAME, (*get name of receipe*)
		eREAD_RECEIPE_NAME_r,
		eWAIT_FOR_COMMAND := 50, (*wait for command of user*)
		eLOAD_RECEIPE, (*SELECT a specific receipe*)
		eLOAD_RECEIPE_r,
		eFETCH_VALUES, (*prepare for read receipe values*)
		eFETCH_VALUES_r,
		eGET_VALUES, (*read each value of receipe*)
		eGET_VALUES_r,
		eSAVE_RECEIPE, (*UPDATE changed values into receipe*)
		eSAVE_RECEIPE_r,
		eSAVE_GET_AFFECTED_ROWS, (*test if saved (if one row is modified)*)
		eSAVE_GET_AFFECTED_ROWS_r,
		eSAVE_AS, (*INSERT changed values into new receipe*)
		eSAVE_AS_r,
		eSAVE_AS_ROWS_AFFECTED, (*test if saved (if one row is modified)*)
		eSAVE_AS_ROWS_AFFECTED_r,
		eDELETE_RECEIPE, (*DELETE receipe*)
		eDELETE_RECEIPE_r,
		eDELETE_ROWS_AFFECTED, (*test if deleted (if one row is modified)*)
		eDELETE_ROWS_AFFECTED_r,
		eRENAME_RECEIPE, (*UPDATE name of receipe*)
		eRENAME_RECEIPE_r,
		eRENAME_GET_AFFECTED_ROWS, (*test if renamed (if one row is modified)*)
		eRENAME_GET_AFFECTED_ROWS_r,
		eDISCONNECT := 150, (*disconnect from server*)
		eDISCONNECT_r,
		eGET_ERROR := 200, (*receive error of server*)
		eGET_ERROR_r,
		eERROR, (*error step*)
		eDUMMY (*dummy step - for development*)
	);
END_TYPE

(*Commands for receipe handling*)

TYPE
	Command_enum :
		(
		eCMD_IDLE, (*nothing to do*)
		eCMD_CONNECT := 10, (*connect to server*)
		eCMD_CONNECT_w,
		eCMD_LOAD := 20, (*load receipe 'sNewReceipe'*)
		eCMD_LOAD_w,
		eCMD_SAVE := 30, (*save receipe 'sActReceipe'*)
		eCMD_SAVE_w,
		eCMD_SAVEAS := 40, (*save as new receipe 'sNewReceipe'*)
		eCMD_SAVEAS_w,
		eCMD_DELETE := 50, (*delete receipe 'sNewReceipe'*)
		eCMD_DELETE_w,
		eCMD_RENAME := 60, (*rename receipe from 'sActReceipe' to 'sNewReceipe'*)
		eCMD_RENAME_w,
		eCMD_DISCONNECT := 70, (*disconnect from server*)
		eCMD_DISCONNECT_w
	);
	CommandInterface_typ : 	STRUCT
		eCommand : Command_enum;
		sActReceipe : STRING[LENGTH_NAME];
		sNewReceipe : STRING[LENGTH_NAME];
		sReceipeNames : ARRAY[0..9] OF STRING[LENGTH_NAME];
		uStatus : UINT; (*0 = OK; 1 = FAIL SQL QUERY; 2 = Unexpected Error*)
		sErrorString : STRING[100];
	END_STRUCT;
END_TYPE
```

#### Variables.var - Local variables
```iecst
(********************************************************************
 * COPYRIGHT --
 ********************************************************************
 * Program: SQLRecipe
 * File: SQLRecipe.var
 * Author: B&R
 * Created: December 27, 2010
 ********************************************************************
 * Local variables of program SQLRecipe
 ********************************************************************)
(*Constants*)
VAR CONSTANT
	LENGTH_NAME : USINT := 30; (*Length of an receipe name*)
END_VAR
(*Configuration Variables*)
VAR
	DBConnectState : dbGetConnState;
	HOST : STRING[40] := '127.0.0.1'; (*Hostname/IP:Port of SQL Server*)
	DATABASE : STRING[40] := 'TestDb'; (*name of database*)
	TABLE : STRING[40] := 'Recipes'; (*name of table*)
	USERNAME : STRING[40] := 'sa'; (*username*)
	PASSWORD : STRING[40] := 'YourStrong@Passw0rd'; (*password*)
END_VAR
(*Variables*)
VAR
	eStep : Steps_enum := (0);
	Command : CommandInterface_typ;
	ConnectionIdent : UDINT := 0;
	sSQLstring : STRING[300] := '';
	ReceipeNameCounter : UDINT := 0;
END_VAR
(*Functionblocks*)
VAR
	ReceipeDBConnect : dbConnect := (0);
	ReceipeDBExecute : dbExecuteSql := (0);
	ReceipeDBErrMsg : dbGetErrorMessage := (0);
	ReceipeDBDisconnect : dbDisconnect := (0);
	ReceipeDBGetData : dbGetData := (0);
	ReceipeDBGetAffectedRows : dbGetAffectedRows := (0);
	ReceipeDBFetchNextRow : dbFetchNextRow := (0);
END_VAR
(*Variables for databaseinterface*)
VAR
	sData : STRING[200] := '';
	usCol : USINT := 0;
END_VAR
```
